TYPE ST_DRIVE_REF : FB_STOEBERSDS_Drive_REF;
END_TYPE

(* stored: Version 1.1.0.1, ProductVersion 3.1.4024.15
   DUT ST_DRIVE_REF: Id {0e37c816-8037-4311-8181-f6f634d3f63d} *)
